(* IEC 61131-3 sources: Test-Git_ESME26/TestProgettoESME_26.fbsproj/TemplateFullProgrammingFramework_Migration.device.xml.v3^/Plc Logic.plclogic.xml.v3^/Application.application.xml.v3^/TemplateFullProgrammingFramework/GlobalVariables, 7 files *)

(* ---- Diagnostics.gvl ---- *)
VAR_GLOBAL
	G_stDiagnosticsToApplicationMarkerarea AT %ML0 : TPL.ST_DiagnosticsToApplicationMarkerArea;
END_VAR

(* ---- ExceptionHandling.gvl ---- *)
VAR_GLOBAL
	G_stExceptionList		: TPL.ST_ExceptionList;
END_VAR

(* ---- HardwareInOuts.gvl ---- *)
VAR_GLOBAL
	G_xMainsContactorOut 		(*-AT %QX0.0-*)	: BOOL;

	G_xEmergencyIn  			(*-AT %IX0.0-*)	: BOOL;
	G_xMainsContactorIn 		(*-AT %IX0.1-*)	: BOOL;
END_VAR

(* ---- InputVariablesEpas.gvl ---- *)
VAR_GLOBAL
	G_xStartEpas				: BOOL;
	G_xStopEpas					: BOOL;
	G_xPrepareEpas				: BOOL;
	G_xAutoEpas					: BOOL;
	G_xHoldEpas					: BOOL;
	G_xAbortEpas				: BOOL;
	G_xProductsOkEpas			: BOOL;
	G_xPowerOnEpas				: BOOL;
	G_xPowerOffEpas				: BOOL;
	G_xManualEpas				: BOOL;
	G_xJogMachineEpas			: BOOL;
	G_xDiagQuitEpas				: BOOL;
	G_xEmergencyEpas			: BOOL := TRUE;
	G_xJogForwEpas				: BOOL;
	G_xJogBackEpas				: BOOL;
	G_xBrakeReleaseEpas			: BOOL;

	G_udiManualModuleSelect		: UDINT;
//	G_udiManualElementSelect	: UDINT;

	G_xDoEnableVis				: BOOL;

	G_xDoPrepare 				: BOOL;
	G_xDoAuto	 				: BOOL;
	G_xDoManual 				: BOOL;
	G_xDoJogMachine 			: BOOL;
	G_xDoBrakeRelease			: BOOL;

	G_xPrepareActive 			: BOOL;
	G_xAutoActive	 			: BOOL;
	G_xManualActive 			: BOOL;
	G_xJogMachineActive 		: BOOL;
	G_xBrakeReleaseActive		: BOOL;
END_VAR

(* ---- InputVariablesExt.gvl ---- *)
VAR_GLOBAL
	G_xStartExt			: BOOL;
	G_xStopExt			: BOOL;
	G_xPrepareExt		: BOOL;
	G_xAutoExt			: BOOL;
	G_xHoldExt			: BOOL;
	G_xAbortExt			: BOOL;
	G_xProductsOkExt	: BOOL;
	G_xPowerOnExt		: BOOL;
	G_xPowerOffExt		: BOOL;
	G_xManualExt		: BOOL;
	G_xJogMachineExt	: BOOL;
	G_xDiagQuitExt		: BOOL;
	G_xJogForwExt		: BOOL;
	G_xJogBackExt		: BOOL;
	G_xBrakeReleaseExt	: BOOL;
END_VAR

(* ---- Logging.gvl ---- *)
VAR_GLOBAL
	G_stLogDataList			: TPL.ST_LogDataList;			(* Global log data list *)
	G_stLogDataListAscii	: TPL.ST_LogDataListAscii;		(* Temp.list for save in XML format *)
	G_stLoggerInterface		: TPL.ST_LoggerInterface;		(* Interface between logger and main machine *)
END_VAR

(* ---- Project.gvl ---- *)
VAR_GLOBAL
	G_diTaskIntervalInMs : DINT;
END_VAR
